(* IEC 61131-3 sources: rusty/tests/lit/single/type_promotion/division, 6 files *)

(* ---- division_guards.st ---- *)
// RUN: %COMPILE %s && %RUN | %CHECK %s
// Divisions and MOD whose result does not depend on the type of the literal.
FUNCTION main : DINT
    VAR
        a : UDINT := 4000000000;
        two : UDINT := 2;
        seven : UDINT := 7;
        ul : ULINT := 18446744073709551615;
        ul2 : ULINT := 2;
        us : USINT := 200;
        ui : UINT := 60000;
        small : UDINT := 100;
        neg : DINT := -7;
        s5 : SINT := 5;
        d2 : DINT := 2;
        ud7 : UDINT := 7;
        q : UDINT;
        ql : ULINT;
        qs : LINT;
        d : DINT;
    END_VAR

    // Two unsigned variables
    q := a / two;
    printf('UDINT 4e9 / UDINT 2 = %u$N', q);                // CHECK: UDINT 4e9 / UDINT 2 = 2000000000
    q := a MOD seven;
    printf('UDINT 4e9 MOD UDINT 7 = %u$N', q);              // CHECK-NEXT: UDINT 4e9 MOD UDINT 7 = 3
    ql := ul / ul2;
    printf('ULINT max / ULINT 2 = %llu$N', ql);             // CHECK-NEXT: ULINT max / ULINT 2 = 9223372036854775807

    // A typed literal of the same type
    q := a / UDINT#2;
    printf('UDINT 4e9 / UDINT#2 = %u$N', q);                // CHECK-NEXT: UDINT 4e9 / UDINT#2 = 2000000000

    // ULINT operands by an untyped literal
    ql := ul / 2;
    printf('ULINT max / 2 = %llu$N', ql);                   // CHECK-NEXT: ULINT max / 2 = 9223372036854775807
    ql := ul MOD 7;
    printf('ULINT max MOD 7 = %llu$N', ql);                 // CHECK-NEXT: ULINT max MOD 7 = 1

    // A literal dividend too large for DINT is LINT
    qs := 4000000000 / two;
    printf('4000000000 / UDINT 2 = %lld$N', qs);            // CHECK-NEXT: 4000000000 / UDINT 2 = 2000000000

    // Values below the signed midpoint
    q := small / 3;
    printf('UDINT 100 / 3 = %u$N', q);                      // CHECK-NEXT: UDINT 100 / 3 = 33
    d := us / 3;
    printf('USINT 200 / 3 = %d$N', d);                      // CHECK-NEXT: USINT 200 / 3 = 66
    d := ui MOD 7;
    printf('UINT 60000 MOD 7 = %d$N', d);                   // CHECK-NEXT: UINT 60000 MOD 7 = 3

    // Signed division cuts towards zero
    d := neg / 2;
    printf('-7 / 2 = %d$N', d);                             // CHECK-NEXT: -7 / 2 = -3
    d := neg MOD 2;
    printf('-7 MOD 2 = %d$N', d);                           // CHECK-NEXT: -7 MOD 2 = -1

    // Mixed signedness and negative literals with non-negative or small operands
    qs := s5 / ul;
    printf('SINT 5 / ULINT max = %lld$N', qs);              // CHECK-NEXT: SINT 5 / ULINT max = 0
    qs := ul / d2;
    printf('ULINT max / DINT 2 = %lld$N', qs);              // CHECK-NEXT: ULINT max / DINT 2 = 9223372036854775807
    qs := ud7 / -2;
    printf('UDINT 7 / -2 = %lld$N', qs);                    // CHECK-NEXT: UDINT 7 / -2 = -3
END_FUNCTION

(* ---- mixed_signedness_variables.st ---- *)
// RUN: %COMPILE %s && %RUN | %CHECK %s
// XFAIL: *
// A signed operand next to a UDINT makes the division signed, and next to a ULINT it makes the division unsigned,
// so one of the two operands is read with the wrong sign.
FUNCTION main : DINT
    VAR
        d5 : DINT := 5;
        sm1 : SINT := -1;
        dm1 : DINT := -1;
        lm1 : LINT := -1;
        s2 : SINT := 2;
        d2 : DINT := 2;
        ul2 : ULINT := 2;
        udmax : UDINT := 4294967295;
        ulmax : ULINT := 18446744073709551615;
        r : LINT;
    END_VAR

    // Signed operand next to a UDINT operand
    r := udmax / d2;
    printf('UDINT max / DINT 2 = %lld$N', r);               // CHECK: UDINT max / DINT 2 = 2147483647
    r := udmax MOD s2;
    printf('UDINT max MOD SINT 2 = %lld$N', r);             // CHECK-NEXT: UDINT max MOD SINT 2 = 1
    r := d5 / udmax;
    printf('DINT 5 / UDINT max = %lld$N', r);               // CHECK-NEXT: DINT 5 / UDINT max = 0

    // Signed operand next to a ULINT operand
    r := dm1 / ul2;
    printf('DINT -1 / ULINT 2 = %lld$N', r);                // CHECK-NEXT: DINT -1 / ULINT 2 = 0
    r := sm1 MOD ul2;
    printf('SINT -1 MOD ULINT 2 = %lld$N', r);              // CHECK-NEXT: SINT -1 MOD ULINT 2 = -1
    r := lm1 / ulmax;
    printf('LINT -1 / ULINT max = %lld$N', r);              // CHECK-NEXT: LINT -1 / ULINT max = 0
END_FUNCTION

(* ---- named_builtin_arguments_with_literal.st ---- *)
// RUN: %COMPILE %s 2> %t.err && %RUN | %CHECK %s
// RUN: not grep -E "Implicit conversion from|Operand of type" %t.err
// An untyped integer literal passed by name to a builtin operator takes the type of the other argument, as
// it does next to the operator, so the operation on a UDINT stays unsigned.
FUNCTION main : DINT
    VAR
        a : UDINT := 4000000000;
        q : UDINT;
    END_VAR

    q := DIV(IN1 := a, IN2 := 2);
    printf('DIV(IN1 := 4e9, IN2 := 2) = %u$N', q);          // CHECK: DIV(IN1 := 4e9, IN2 := 2) = 2000000000
    q := DIV(IN2 := 2, IN1 := a);
    printf('DIV(IN2 := 2, IN1 := 4e9) = %u$N', q);          // CHECK-NEXT: DIV(IN2 := 2, IN1 := 4e9) = 2000000000
    q := MOD(IN1 := a, IN2 := 7);
    printf('MOD(IN1 := 4e9, IN2 := 7) = %u$N', q);          // CHECK-NEXT: MOD(IN1 := 4e9, IN2 := 7) = 3
    q := SUB(IN1 := a, IN2 := 1);
    printf('SUB(IN1 := 4e9, IN2 := 1) = %u$N', q);          // CHECK-NEXT: SUB(IN1 := 4e9, IN2 := 1) = 3999999999
    q := a / 2;
    printf('4e9 / 2 = %u$N', q);                            // CHECK-NEXT: 4e9 / 2 = 2000000000
END_FUNCTION

(* ---- udint_by_untyped_literal.st ---- *)
// RUN: %COMPILE %s && %RUN | %CHECK %s
// An untyped integer literal takes the type of a UDINT operand, so the division is unsigned.
FUNCTION main : DINT
    VAR
        a : UDINT := 4000000000;
        q : UDINT;
    END_VAR

    q := a / 2;
    printf('UDINT 4e9 / 2 = %u$N', q);                      // CHECK: UDINT 4e9 / 2 = 2000000000
    q := a / 3;
    printf('UDINT 4e9 / 3 = %u$N', q);                      // CHECK-NEXT: UDINT 4e9 / 3 = 1333333333
    q := a / 2147483647;
    printf('UDINT 4e9 / 2147483647 = %u$N', q);             // CHECK-NEXT: UDINT 4e9 / 2147483647 = 1
    q := a MOD 7;
    printf('UDINT 4e9 MOD 7 = %u$N', q);                    // CHECK-NEXT: UDINT 4e9 MOD 7 = 3
    q := a MOD 2147483647;
    printf('UDINT 4e9 MOD 2147483647 = %u$N', q);           // CHECK-NEXT: UDINT 4e9 MOD 2147483647 = 1852516353
    q := (a / 2) MOD 7;
    printf('(UDINT 4e9 / 2) MOD 7 = %u$N', q);              // CHECK-NEXT: (UDINT 4e9 / 2) MOD 7 = 5
END_FUNCTION

(* ---- unsigned_by_negative_literal.st ---- *)
// RUN: %COMPILE %s && %RUN | %CHECK %s
// XFAIL: *
// A negative literal next to a UDINT makes the division signed in 32 bits, and next to a ULINT it is read as unsigned.
FUNCTION main : DINT
    VAR
        udmax : UDINT := 4294967295;
        ul5 : ULINT := 5;
        r : LINT;
    END_VAR

    // UDINT dividend
    r := udmax / -2;
    printf('UDINT max / -2 = %lld$N', r);                   // CHECK: UDINT max / -2 = -2147483647
    r := udmax MOD -2;
    printf('UDINT max MOD -2 = %lld$N', r);                 // CHECK-NEXT: UDINT max MOD -2 = 1

    // ULINT dividend
    r := ul5 / -2;
    printf('ULINT 5 / -2 = %lld$N', r);                     // CHECK-NEXT: ULINT 5 / -2 = -2
END_FUNCTION

(* ---- literal_by_declaration_section.st ---- *)
// RUN: %COMPILE %s && %RUN | %CHECK %s
// A UDINT operand divided by an untyped literal stays UDINT, wherever the operand is declared.
VAR_GLOBAL
    g : UDINT := 4294967295;
END_VAR

VAR_GLOBAL CONSTANT
    gc : UDINT := 4294967295;
END_VAR

FUNCTION_BLOCK probe
    VAR_INPUT
        i : UDINT;
    END_VAR
    VAR_INPUT CONSTANT
        ic : UDINT := 4294967295;
    END_VAR
    VAR_IN_OUT
        io : UDINT;
    END_VAR
    VAR_OUTPUT
        o : UDINT;
    END_VAR
    VAR CONSTANT
        c : UDINT := 4294967295;
    END_VAR
    VAR_TEMP
        t : UDINT;
    END_VAR
    VAR
        q : ULINT;
    END_VAR

    o := 4294967295;
    t := 4294967295;
    q := i / 2;
    printf('VAR_INPUT / 2 = %llu$N', q);
    q := ic MOD 7;
    printf('VAR_INPUT CONSTANT MOD 7 = %llu$N', q);
    q := io / 2;
    printf('VAR_IN_OUT / 2 = %llu$N', q);
    q := io MOD 7;
    printf('VAR_IN_OUT MOD 7 = %llu$N', q);
    q := o / 2;
    printf('VAR_OUTPUT / 2 = %llu$N', q);
    q := c MOD 7;
    printf('VAR CONSTANT MOD 7 = %llu$N', q);
    q := t / 2;
    printf('VAR_TEMP / 2 = %llu$N', q);
    q := g MOD 7;
    printf('VAR_GLOBAL MOD 7 = %llu$N', q);
    q := gc / 2;
    printf('VAR_GLOBAL CONSTANT / 2 = %llu$N', q);
END_FUNCTION_BLOCK

FUNCTION main : DINT
    VAR
        inst : probe;
        v : UDINT := 4294967295;
    END_VAR

    inst(i := 4294967295, io := v);
    // CHECK: VAR_INPUT / 2 = 2147483647
    // CHECK-NEXT: VAR_INPUT CONSTANT MOD 7 = 3
    // CHECK-NEXT: VAR_IN_OUT / 2 = 2147483647
    // CHECK-NEXT: VAR_IN_OUT MOD 7 = 3
    // CHECK-NEXT: VAR_OUTPUT / 2 = 2147483647
    // CHECK-NEXT: VAR CONSTANT MOD 7 = 3
    // CHECK-NEXT: VAR_TEMP / 2 = 2147483647
    // CHECK-NEXT: VAR_GLOBAL MOD 7 = 3
    // CHECK-NEXT: VAR_GLOBAL CONSTANT / 2 = 2147483647
END_FUNCTION
